FUNCTION_BLOCK MOD_StateGate (* The module's front desk inside MOD_StateManager: answers Reset, Start, Stop, Abort or Clear at once (only from the module's owner, only in a state PackML allows it in) and passes an accepted command on to MOD_StateLogic. Technical: Decides the module commands Reset/Start/Stop/Abort/Clear: only from the occupation owner (5 NotPermitted) and only in a state PackML allows them in (4 NotReady); passes an accepted one on to MOD_StateLogic *)
  (* Standard: 61499-2 *)
  (* Version 0.1, 2026-09-28, Project contributors, AAU Smart Production Lab *)
  PACKAGE modlib;
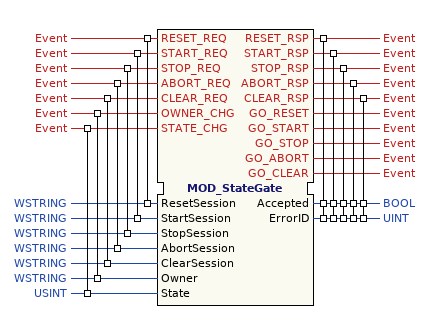
  EVENT_INPUT
    RESET_REQ WITH ResetSession; (* RESET(Session) was called *)
    START_REQ WITH StartSession; (* START(Session) was called *)
    STOP_REQ WITH StopSession; (* STOP(Session) was called *)
    ABORT_REQ WITH AbortSession; (* ABORT(Session) was called *)
    CLEAR_REQ WITH ClearSession; (* CLEAR(Session) was called *)
    OWNER_CHG WITH Owner; (* The owner changed *)
    STATE_CHG WITH State; (* The module's state changed (State, as MOD_StateLogic publishes it) *)
  END_EVENT
  EVENT_OUTPUT
    RESET_RSP WITH Accepted, ErrorID; (* Answer to RESET: Accepted, ErrorID *)
    START_RSP WITH Accepted, ErrorID; (* Answer to START: Accepted, ErrorID *)
    STOP_RSP WITH Accepted, ErrorID; (* Answer to STOP: Accepted, ErrorID *)
    ABORT_RSP WITH Accepted, ErrorID; (* Answer to ABORT: Accepted, ErrorID *)
    CLEAR_RSP WITH Accepted, ErrorID; (* Answer to CLEAR: Accepted, ErrorID *)
    GO_RESET; (* Reset the module: an accepted Reset(Session) *)
    GO_START; (* Start the module: an accepted Start(Session) *)
    GO_STOP; (* Stop the module: an accepted Stop(Session) *)
    GO_ABORT; (* Abort the module: an accepted Abort(Session) *)
    GO_CLEAR; (* Clear the module: an accepted Clear(Session) *)
  END_EVENT
  VAR_INPUT
    ResetSession : WSTRING; (* Session ID of the caller of Reset *)
    StartSession : WSTRING; (* Session ID of the caller of Start *)
    StopSession : WSTRING; (* Session ID of the caller of Stop *)
    AbortSession : WSTRING; (* Session ID of the caller of Abort *)
    ClearSession : WSTRING; (* Session ID of the caller of Clear *)
    Owner : WSTRING; (* Session ID of the module's owner (empty: free) *)
    State : USINT := 2; (* PackML state: 1 Clearing, 2 Stopped, 3 Starting, 4 Idle, 6 Execute, 7 Stopping, 8 Aborting, 9 Aborted, 15 Resetting *)
  END_VAR
  VAR_OUTPUT
    Accepted : BOOL; (* The call was accepted *)
    ErrorID : UINT; (* Error code: 0 none, 1 PreconditionViolated, 2 InvariantViolated, 3 Timeout, 4 NotReady, 5 NotPermitted, 6 Busy, 7 Interrupted, 8 OutOfRange *)
  END_VAR
  VAR
    Owned : BOOL;
  END_VAR
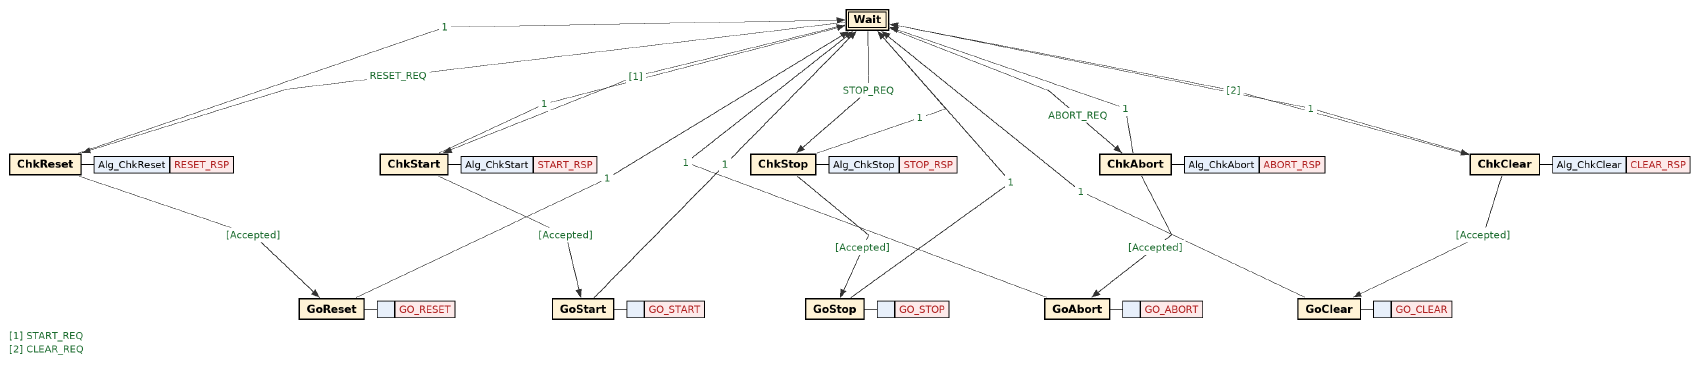
  EC_STATES
    Wait;
    ChkReset : Alg_ChkReset -> RESET_RSP;
    GoReset : -> GO_RESET;
    ChkStart : Alg_ChkStart -> START_RSP;
    GoStart : -> GO_START;
    ChkStop : Alg_ChkStop -> STOP_RSP;
    GoStop : -> GO_STOP;
    ChkAbort : Alg_ChkAbort -> ABORT_RSP;
    GoAbort : -> GO_ABORT;
    ChkClear : Alg_ChkClear -> CLEAR_RSP;
    GoClear : -> GO_CLEAR;
  END_STATES
  EC_TRANSITIONS
    Wait TO ChkReset := RESET_REQ;
    ChkReset TO GoReset := [Accepted];
    ChkReset TO Wait := 1;
    GoReset TO Wait := 1;
    Wait TO ChkStart := START_REQ;
    ChkStart TO GoStart := [Accepted];
    ChkStart TO Wait := 1;
    GoStart TO Wait := 1;
    Wait TO ChkStop := STOP_REQ;
    ChkStop TO GoStop := [Accepted];
    ChkStop TO Wait := 1;
    GoStop TO Wait := 1;
    Wait TO ChkAbort := ABORT_REQ;
    ChkAbort TO GoAbort := [Accepted];
    ChkAbort TO Wait := 1;
    GoAbort TO Wait := 1;
    Wait TO ChkClear := CLEAR_REQ;
    ChkClear TO GoClear := [Accepted];
    ChkClear TO Wait := 1;
    GoClear TO Wait := 1;
  END_TRANSITIONS
  ALGORITHM Alg_ChkReset IN ST:
Owned := (ResetSession = Owner) AND (Owner <> "");
Accepted := Owned AND ((State = 2));
IF NOT Owned THEN
  ErrorID := 5;
ELSIF NOT Accepted THEN
  ErrorID := 4;
ELSE
  ErrorID := 0;
END_IF;
  END_ALGORITHM
  ALGORITHM Alg_ChkStart IN ST:
Owned := (StartSession = Owner) AND (Owner <> "");
Accepted := Owned AND ((State = 4));
IF NOT Owned THEN
  ErrorID := 5;
ELSIF NOT Accepted THEN
  ErrorID := 4;
ELSE
  ErrorID := 0;
END_IF;
  END_ALGORITHM
  ALGORITHM Alg_ChkStop IN ST:
Owned := (StopSession = Owner) AND (Owner <> "");
Accepted := Owned AND ((State = 4) OR (State = 6) OR (State = 15));
IF NOT Owned THEN
  ErrorID := 5;
ELSIF NOT Accepted THEN
  ErrorID := 4;
ELSE
  ErrorID := 0;
END_IF;
  END_ALGORITHM
  ALGORITHM Alg_ChkAbort IN ST:
Owned := (AbortSession = Owner) AND (Owner <> "");
Accepted := Owned AND ((State = 2) OR (State = 4) OR (State = 6) OR (State = 7) OR (State = 15));
IF NOT Owned THEN
  ErrorID := 5;
ELSIF NOT Accepted THEN
  ErrorID := 4;
ELSE
  ErrorID := 0;
END_IF;
  END_ALGORITHM
  ALGORITHM Alg_ChkClear IN ST:
Owned := (ClearSession = Owner) AND (Owner <> "");
Accepted := Owned AND ((State = 9));
IF NOT Owned THEN
  ErrorID := 5;
ELSIF NOT Accepted THEN
  ErrorID := 4;
ELSE
  ErrorID := 0;
END_IF;
  END_ALGORITHM
END_FUNCTION_BLOCK
